Fanuc KAREL source: KT00831.KL

PROGRAM KT00831
%NOLOCKGROUP
VAR
  S1: STRING[80]
  S2: STRING[80]
  OUT: REAL
BEGIN
  S1 = 'A'
  S2 = 'B'
  S1 = 'A'
  S2 = 'B'
  OUT = SIN(S1)
END KT00831
